PROGRAM main
  VAR
    Button AT %QX0.0 : BOOL;
    Motor AT %QX0.1 : BOOL;
    Package_sense AT %QX0.2 : BOOL;
    reset_counter AT %QX0.3 : BOOL;
    total_count AT %MW1 : INT;
    CTU0 : CTU;
  END_VAR

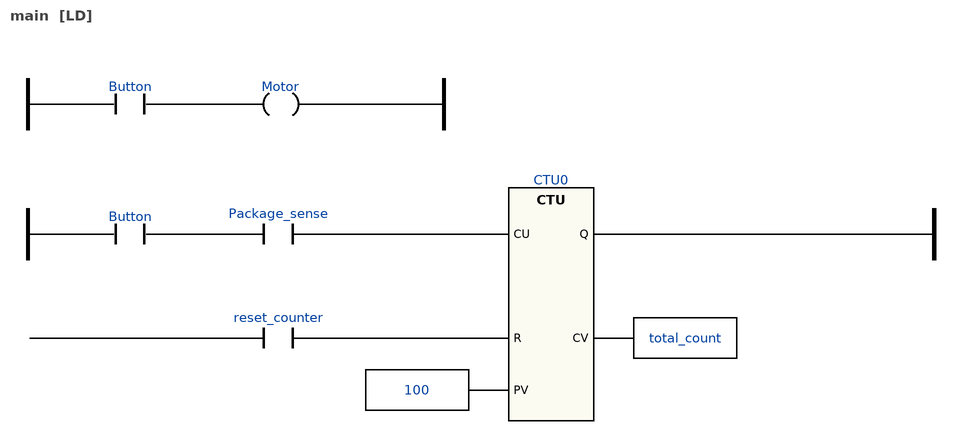
(* LD diagram, written out as Structured Text *)
Motor := Button;
CTU0(CU := Button AND Package_sense, R := reset_counter, PV := 100);
total_count := CTU0.CV;
END_PROGRAM
